Staubli VAL3: onStart.pgx

public program onStart()
  local num l_i
begin
  //list
  resize(sActionList,1,size(actdata:aActItem))
  for l_i = 0 to size(sActionList)-1
    sActionList[l_i]=toString("",l_i)+","+actdata:aActItem[l_i].sComment
  endFor
  //
  //  resize(sIOList,1,size(io:dInItem))
  //  for l_i = 0 to size(sIOList)-1
  //    sIOList[l_i]=toString("",l_i)
  //  endFor
  //  //
  insert(sActionList[0])
  sActionList[0]="--"
  //insert(sIOList[0])
  sLastList=""
  sSelIO="--"
end
